(* IEC 61131-3 sources: rusty/tests/lit/multi/duplicate_symbol_fb_output_and_enum, 1 file *)

(* ---- main.st ---- *)
PROGRAM mainProg
VAR
    fb : MC_ReadStatus;
END_VAR
    fb();

    printf('%d$N', fb.StatusEnumerator);
    printf('%d$N', fb.Homing);
END_PROGRAM

FUNCTION main
    mainProg();
END_FUNCTION
